// TIA Portal V19 export
DATA_BLOCK "GVL"   // DB2
{ S7_Optimized_Access := 'TRUE' }
// stored: MemoryReserve 100
   VAR
      xKillAll : Bool;
      xSystemWakeUp : Bool;
      Auto : Bool;
      Manual : Bool;
      Servo : "ST_Servo";
      ExitConveyor_Start : Bool;
      Robot { S7_SetPoint := 'True'} : Array[1..3] of "ST_ROBOT";
      PickPosition { S7_SetPoint := 'True'} : "ST_PICK_POSITION";
      PlacePosition { S7_SetPoint := 'True'} : "ST_PLACE_POSITION";
      Place_Empty { S7_SetPoint := 'True'} : "ST_Pos";
      SystemWakeUp { S7_SetPoint := 'True'} : Bool;
      xAttemptKillAll : Bool;
      xBlink : Bool;
      xBlinkFast : Bool;
      Global_ms : UDInt;
      xTick100ms : Bool;
      mm : Bool;
      EnableTest : Bool;
      xSystemStart : Bool;
      xCommissioning : Bool;
   END_VAR
BEGIN
END_DATA_BLOCK
